FUNCTION_BLOCK F (* Negative C3: REQ guards read the position from a carried-over variable *)
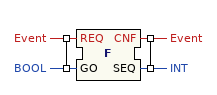
  EVENT_INPUT
    REQ WITH GO;
  END_EVENT
  EVENT_OUTPUT
    CNF WITH SEQ;
  END_EVENT
  VAR_INPUT
    GO : BOOL;
  END_VAR
  VAR_OUTPUT
    SEQ : INT;
  END_VAR
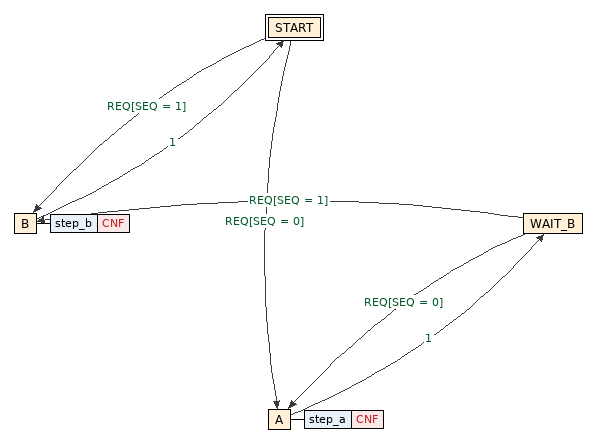
  EC_STATES
    START;
    WAIT_B;
    A : step_a -> CNF;
    B : step_b -> CNF;
  END_STATES
  EC_TRANSITIONS
    START TO A := REQ[SEQ = 0];
    START TO B := REQ[SEQ = 1];
    WAIT_B TO A := REQ[SEQ = 0];
    WAIT_B TO B := REQ[SEQ = 1];
    A TO WAIT_B := 1;
    B TO START := 1;
  END_TRANSITIONS
  ALGORITHM step_a IN ST:
SEQ := 0;
IF GO THEN
  SEQ := 1;
END_IF;
  END_ALGORITHM
  ALGORITHM step_b IN ST:
IF NOT GO THEN
  SEQ := 0;
END_IF;
  END_ALGORITHM
END_FUNCTION_BLOCK
